(* IEC 61131-3 sources: rung/tests/conformance/cases/support, 4 files *)

(* ---- E_ConformanceState.st ---- *)
(* SPDX-License-Identifier: MIT *)
TYPE E_ConformanceState :
(
    Idle := 0,
    Running := 10,
    Stopping := 11
) INT := Idle;
END_TYPE

(* ---- ST_ConformancePair.st ---- *)
(* SPDX-License-Identifier: MIT *)
TYPE ST_ConformancePair :
STRUCT
    number : INT;
    flag : BOOL;
END_STRUCT
END_TYPE

(* ---- FC_ConformanceReturn.st ---- *)
(* SPDX-License-Identifier: MIT *)
FUNCTION FC_ConformanceReturn : INT
VAR_INPUT
    value : INT;
END_VAR
FC_ConformanceReturn := value;
IF value < 0 THEN
    RETURN;
END_IF
FC_ConformanceReturn := value + 10;
END_FUNCTION

(* ---- FB_ConformanceAccumulate.st ---- *)
(* SPDX-License-Identifier: MIT *)
FUNCTION_BLOCK FB_ConformanceAccumulate
VAR_INPUT
    increment : INT;
END_VAR
VAR_OUTPUT
    total : INT;
END_VAR
total := total + increment;
END_FUNCTION_BLOCK
